Fanuc KAREL source: ka00054.KL

PROGRAM KA00054
%STACKSIZE=65535
%PRIORITY=65535
%NOLOCKGROUP
VAR
SRC : POSITION
DST : XYZWPR
BEGIN
DST=SRC
END KA00054
